Staubli VAL3: Point2Trsf.pgx

public program Point2Trsf(point x_pPoint, trsf& x_trTrsf)
begin
  x_trTrsf.x=x_pPoint.trsf.x
  x_trTrsf.y=x_pPoint.trsf.y
  x_trTrsf.z=x_pPoint.trsf.z
  x_trTrsf.rx=x_pPoint.trsf.rx
  x_trTrsf.ry=x_pPoint.trsf.ry
  x_trTrsf.rz=x_pPoint.trsf.rz
end
